FUNCTION_BLOCK FB_InstrumentationScope
VAR_OUTPUT
	name: T_MaxString;
	version: T_MaxString;
	droppedAttributesCount: UDINT;
	schemaUrl: T_MaxString;
END_VAR
VAR_OUTPUT
	attributes: FB_Attributes(maxCount := TcOtlp_GVL.DEFAULT_MAX_ATTRIBUTE_COUNT);
END_VAR

METHOD copyFrom : BOOL
VAR_IN_OUT
	src: FB_InstrumentationScope;
END_VAR
VAR_OUTPUT
	failureResult: E_AttributesFailureReason;
END_VAR
failureResult := E_AttributesFailureReason.NA;
THIS^.name := src.name;
THIS^.version := src.version;
THIS^.droppedAttributesCount := src.droppedAttributesCount;
THIS^.schemaUrl := src.schemaUrl;
THIS^.attributes.free();
copyFrom := THIS^.attributes.copyFrom(src:=src.attributes, failureReason=>failureResult);
END_METHOD

//FB_Exit must be implemented explicitly. If there is an implementation, then the
//method is called before the controller removes the code of the function block instance
//(implicit call). The return value is not evaluated.
METHOD FB_Exit: BOOL
VAR_INPUT
    bInCopyCode: BOOL;  // TRUE: the exit method is called in order to leave the instance which will be copied afterwards (online change).  
END_VAR
THIS^.free();
END_METHOD

METHOD FB_Init: BOOL
VAR_INPUT
	bInitRetains: BOOL;
	bInCopyCode: BOOL;
	name: T_MaxString;
	version: T_MaxString;
	schemaUrl: T_MaxString;
END_VAR
THIS^.name := name;
THIS^.version := version;
THIS^.schemaUrl := schemaUrl;
END_METHOD

METHOD free
VAR_INPUT
END_VAR
THIS^.attributes.free();
END_METHOD

END_FUNCTION_BLOCK

(* stored: Version 1.1.0.1
   POU FB_InstrumentationScope: Id {b7d10966-7b60-4f22-b7d9-720144dd9472}, SpecialFunc None
   Method copyFrom: Id {545489b4-e9b6-45f4-bd71-13b12b5d895a}
   Method FB_Exit: Id {dfd2f978-3108-4426-a903-5c90d7c5bec7}
   Method FB_Init: Id {f1944aeb-9f9c-4684-855f-98ad767fb9b0}
   Method free: Id {b8940d1a-768c-4234-9b2f-4caa954f371f} *)
